Yaskawa INFORM job: TURNPRO.JBI

/JOB
//NAME TURNPRO
//POS
///NPOS 9,0,0,0,0,0
///TOOL 9
///POSTYPE PULSE
///PULSE
C00000=204800,0,0,-34475,0,0,0
C00001=0,0,229831,-34475,0,0,0
C00002=0,0,0,-34475,-229831,0,0
C00003=-204800,0,0,-34475,229831,0,0
C00004=0,194560,0,-218340,0,-110251,-218340
C00005=-92160,-30720,-206848,34475,206848,0,68949
C00006=358400,0,402204,-34475,-620544,203093,0
C00007=-184320,0,-206848,0,620544,-104448,0
C00008=358400,0,402204,-34475,-620544,203093,0
//INST
<volatile>
///COMM Generated using RoboDK
///ATTR SC,RW
///GROUP1 RB1
NOP
'Program generated by RoboDK v
'6.0.7 for Yaskawa Motoman CSD
'A10F on XX/XX/XXXX 18:00:00
'Using nominal kinematics.
'Using Frame S (targets wrt ba
'se):
'1234.6,-98.8,50.5,0.0,0.0,30.
'0
'Tool Tool S should be close t
'o:
'10.0,20.0,150.0,0.0,0.0,0.0
MOVL C00000 V=100.0
MOVL C00001 V=100.0
MOVL C00002 V=100.0
MOVL C00003 V=100.0
MOVL C00004 V=100.0
MOVL C00005 V=100.0
MOVL C00006 V=100.0
MOVL C00007 V=100.0
MOVJ C00008 VJ=50.00
END
